// TIA Portal V20 export
DATA_BLOCK "HMI_BETR_ART_POS"   // DB2003
{ S7_Optimized_Access := 'FALSE' }
// stored: AutoNumber false
   VAR
      POS3_0 { S7_SetPoint := 'True'} : "WinCC_Stationsvariablen";
      POS3_1 { S7_SetPoint := 'True'} : "WinCC_Stationsvariablen";
      POS3_2 { S7_SetPoint := 'True'} : "WinCC_Stationsvariablen";
      POS3_3 { S7_SetPoint := 'True'} : "WinCC_Stationsvariablen";
      POS3_4 { S7_SetPoint := 'True'} : "WinCC_Stationsvariablen";
      POS4_0 { S7_SetPoint := 'True'} : "WinCC_Stationsvariablen";
      POS4_0_Zuführung { S7_SetPoint := 'True'} : "WinCC_Stationsvariablen";
      POS5_0 { S7_SetPoint := 'True'} : "WinCC_Stationsvariablen";
      POS5_0_Zuführung { S7_SetPoint := 'True'} : "WinCC_Stationsvariablen";
      POS6_0 { S7_SetPoint := 'True'} : "WinCC_Stationsvariablen";
      POS7_0 { S7_SetPoint := 'True'} : "WinCC_Stationsvariablen";
      POS7_1 { S7_SetPoint := 'True'} : "WinCC_Stationsvariablen";
      POS7_2 { S7_SetPoint := 'True'} : "WinCC_Stationsvariablen";
      POS7_3 { S7_SetPoint := 'True'} : "WinCC_Stationsvariablen";
      POS7_4 { S7_SetPoint := 'True'} : "WinCC_Stationsvariablen";
      POS8_0 { S7_SetPoint := 'True'} : "WinCC_Stationsvariablen";
      POS8_1 { S7_SetPoint := 'True'} : "WinCC_Stationsvariablen";
      POS8_2 { S7_SetPoint := 'True'} : "WinCC_Stationsvariablen";
      POS8_3 { S7_SetPoint := 'True'} : "WinCC_Stationsvariablen";
      POS9_0 { S7_SetPoint := 'True'} : "WinCC_Stationsvariablen";
      POS9_1 { S7_SetPoint := 'True'} : "WinCC_Stationsvariablen";
      POS9_2 { S7_SetPoint := 'True'} : "WinCC_Stationsvariablen";
      POS9_3 { S7_SetPoint := 'True'} : "WinCC_Stationsvariablen";
      POS9_4 { S7_SetPoint := 'True'} : "WinCC_Stationsvariablen";
      POS9_5 { S7_SetPoint := 'True'} : "WinCC_Stationsvariablen";
      POS9_6 { S7_SetPoint := 'True'} : "WinCC_Stationsvariablen";
      POS10_0 { S7_SetPoint := 'True'} : "WinCC_Stationsvariablen";
      POS11 { S7_SetPoint := 'True'} : "WinCC_Stationsvariablen";
      POS12 { S7_SetPoint := 'True'} : "WinCC_Stationsvariablen";
   END_VAR
BEGIN
END_DATA_BLOCK
